KUKA KRL program: main_lab.src

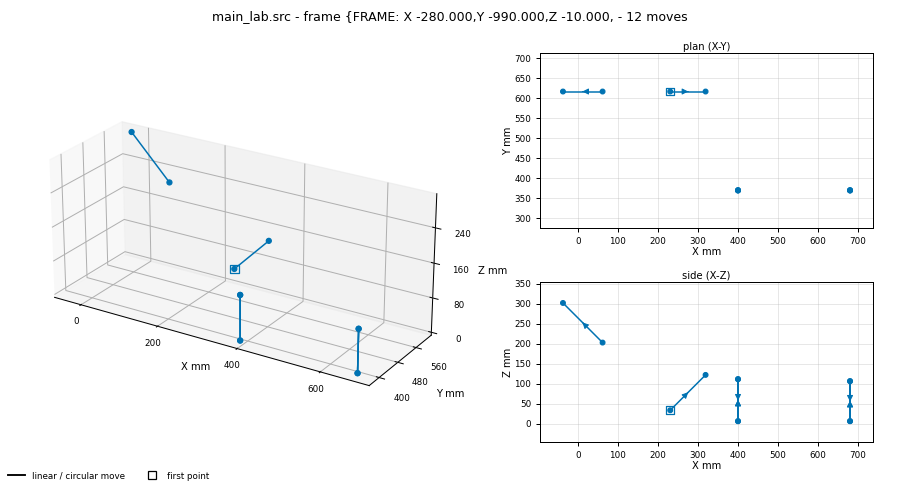
[picture p0: tool path of main_lab.src in frame {FRAME: X -280.000,Y -990.000,Z -10.000,, 12 of 19 moves have a stored position in this frame; points joined in program order, loops and branches not executed]
&ACCESS RVP
&REL 1
&PARAM TEMPLATE = C:\KRC\Roboter\Template\vorgabe
&PARAM EDITMASK = *
DEF main_lab ( )


EXT BAS (BAS_COMMAND :IN,REAL :IN )


; GLOBAL INTERRUPT DECL 3 WHEN $STOPMESS==TRUE DO IR_STOPM ( )
; INTERRUPT ON 3

;FOLD Initialise and set default speed
BAS (#INITMOV,0)
BAS (#VEL_PTP,10)   ; Laborvorgabe: PTP 10 %
BAS (#ACC_PTP,20)
$VEL.CP=0.05        ; 50 mm/s (Laborvorgabe reduziert: 0.005 m/s) - Override am Pendant zusaetzlich niedrig halten
BAS (#TOOL,0)
BAS (#BASE,0)
;ENDFOLD

;;FOLD STARTPOS
;$BWDSTART = FALSE
;PDAT_ACT = PDEFAULT
;BAS(#PTP_DAT)
;FDAT_ACT = {TOOL_NO 0,BASE_NO 0,IPO_FRAME #BASE}
;BAS(#FRAMES)
;;ENDFOLD

$ADVANCE = 5

;FOLD ---- Quickly skip BCO ----
; PTP $AXIS_ACT
;ENDFOLD

;FOLD ---- GO HOME ----
; PTP {A1 0.000, A2 -90.000, A3 90.000, A4 0.000, A5 0.000, A6 0.000, E1 0, E2 0, E3 0, E4 0, E5 0, E6 0}
;ENDFOLD


; Laborversion: Greifer ueber $OUT[5]/$OUT[6], factory_reset entfernt
; Program generated by RoboDK v6.0.7 for KUKA KR 6 R900 sixx on 07/11/2026 19:20:57
; Using nominal kinematics.
; ---- Laborausstattung initialisieren ----
$ANOUT[3] = 0.15    ; Druck Kollisionserkennung
; ---- Greifer oeffnen ----
$OUT[6] = FALSE
$OUT[5] = TRUE
WAIT SEC 1
; ---- Setting reference (Base) ----
$BASE = {FRAME: X -280.000,Y -990.000,Z -10.000,A 0.000,B 0.000,C 0.000}
; --------------------------
; ---- Setting tool (TCP) ----
$TOOL = {FRAME: X 0.000,Y 0.000,Z 288.000,A 43.000,B 0.000,C 0.000}
; --------------------------
PTP {A1 90.00000,A2 -90.00000,A3 90.00000,A4 0.00000,A5 90.00000,A6 0.00000}
; ---- Greifer oeffnen ----
$OUT[6] = FALSE
$OUT[5] = TRUE
WAIT SEC 1
PTP {A1 51.26700,A2 -51.81700,A3 122.51100,A4 40.26010,A5 58.59630,A6 -119.41200}
LIN {X 230.579,Y 617.000,Z 34.236,A 0.000,B 45.000,C 180.000}
; ---- Greifer schliessen ----
$OUT[5] = FALSE
$OUT[6] = TRUE
WAIT SEC 1
; Attach to gripper_TCP
LIN {X 318.967,Y 617.000,Z 122.624,A 0.000,B 45.000,C -180.000}
PTP {A1 79.04590,A2 -50.21190,A3 96.54170,A4 0.00000,A5 43.67020,A6 -57.95410}
LIN {X 400.000,Y 370.000,Z 7.000,A 0.000,B 0.000,C -180.000}
; ---- Greifer oeffnen ----
$OUT[6] = FALSE
$OUT[5] = TRUE
WAIT SEC 1
; Detach from gripper_TCP
LIN {X 400.000,Y 370.000,Z 112.000,A 0.000,B 0.000,C 180.000}
LIN {X 400.000,Y 370.000,Z 7.000,A 0.000,B 0.000,C -180.000}
; ---- Greifer schliessen ----
$OUT[5] = FALSE
$OUT[6] = TRUE
WAIT SEC 1
; Attach to gripper_TCP
LIN {X 400.000,Y 370.000,Z 112.000,A 0.000,B 0.000,C 180.000}
PTP {A1 57.17150,A2 -38.93430,A3 75.31350,A4 0.00000,A5 53.62070,A6 -169.82900}
LIN {X 680.000,Y 370.000,Z 7.000,A -90.000,B 0.000,C -180.000}
; ---- Greifer oeffnen ----
$OUT[6] = FALSE
$OUT[5] = TRUE
WAIT SEC 1
; Detach from gripper_TCP
LIN {X 680.000,Y 370.000,Z 107.000,A -90.000,B 0.000,C 180.000}
LIN {X 680.000,Y 370.000,Z 7.000,A -90.000,B 0.000,C -180.000}
; ---- Greifer schliessen ----
$OUT[5] = FALSE
$OUT[6] = TRUE
WAIT SEC 1
; Attach to gripper_TCP
LIN {X 680.000,Y 370.000,Z 107.000,A -90.000,B 0.000,C 180.000}
PTP {A1 90.00000,A2 -90.00000,A3 90.00000,A4 0.00000,A5 90.00000,A6 0.00000}
PTP {A1 98.72560,A2 -83.01650,A3 132.96600,A4 61.91930,A5 52.38900,A6 -83.59410}
LIN {X 61.532,Y 617.000,Z 203.436,A 0.000,B 45.000,C -180.000}
; ---- Greifer oeffnen ----
$OUT[6] = FALSE
$OUT[5] = TRUE
WAIT SEC 1
; Detach from gripper_TCP
LIN {X -37.463,Y 617.000,Z 302.431,A 0.000,B 45.000,C -180.000}
PTP {A1 90.00000,A2 -90.00000,A3 90.00000,A4 0.00000,A5 90.00000,A6 0.00000}
END
